Fanuc KAREL source: KB00014.KL

PROGRAM KB00014
%NOLOCKGROUP
%ENVIRONMENT FLBT
VAR
  P1: FILE
  RESULT: INTEGER
BEGIN
  RESULT = BYTES_LEFT(P1)
END KB00014
